{attribute 'qualified_only'}

VAR_GLOBAL
	Shutter1MorningScheduler : fbScheduler;
	Shutter1EveningScheduler : fbScheduler;


															
															
END_VAR

(* stored: Version 1.1.0.1
   GVL gvlScheduler: Id {f0dfc590-e34c-421b-b16b-08f06907ee9a} *)
